Fanuc KAREL source: KT00490.KL

PROGRAM KT00490
%NOLOCKGROUP
VAR
  P1: POSITION
  P2: JOINTPOS
  OUT: XYZWPR
BEGIN
  OUT = P1 : P2
END KT00490
